// TIA Portal V19 export
TYPE "EM02_Input"
   STRUCT
      Cmds { S7_SetPoint := 'True'} : "EM_Input";
      CtrlMode : Int;   // 0=Off, 1=PID local, 2=PID externo (SeedMaster), 3=Ruptura de vacÃ­o
      VaccumSP : Real;   // Setpoint en mbar para control Local
      AtmPressure : Real := 1013.25;   // PresiÃ³n atmosfÃ©rica en mbar
      VaccumValid : Bool := TRUE;
      VaccumFilter : Time := T#3S;
      VaccumBand : Real := 10.0;   // Banda de validez alrededor del SP en mbar (|PV - SP| <= banda)
      VaccumTimeout : Time;
      VaccumSMMV : Real;   // Variable manipulada externa en porcentaje, rango 0..100
   END_STRUCT;
END_TYPE
